(* Release Left Axis *)
IF _SubStep.isActive(2) THEN 
	axis1.Enable:= TRUE;
	IF NOT axis1.State.finish THEN 
		_updateHmiTextWithAxisBusy(axisName:= axisName1);
	ELSIF NOT axis1.State.pass THEN 
		_addressRestart:= _SubStep.actual;
		_subStepError:= "Left axis in error";;
		_subStepMessage:= axis1.State.description;
		_SubStep.set(request:= _SUB_ADDRESS_RETRY_ABORT);
	ELSE 
		_SubStep.INC();
	END_IF
END_IF
(* Reset Axis Right *)
IF _SubStep.isActive(3) THEN 
	IF axis2.Fault THEN 
	axis2.ResetFault();
		IF NOT axis2.AxisError THEN 
			_SubStep.INC();
		ELSE 
			_updateHmiTextWithAxisBusy(axisName:= axisName2); 
		END_IF
	ELSE 
		_SubStep.INC();
	END_IF
END_IF

(* Enable Axis Right *)
IF _SubStep.isActive(4) THEN 
	axis2.Ex_On();
	IF NOT axis2.State.finish THEN 
		_updateHmiTextWithAxisBusy(axisName:= axisName2);
	ELSIF NOT axis2.State.pass THEN 
		_subStepError:= "Right axis in error";
		_subStepMessage:= axis2.State.description;
		_SubStep.set(request:= _SUB_ADDRESS_RETRY_ABORT);
	ELSIF axis2.AxisIsOn THEN 
		_SubStep.INC();
	ELSE 
		_updateHmiTextWithAxisBusy(axisName:= axisName2);
	END_IF
END_IF

(* Release Axis Right *)
IF _SubStep.isActive(5) THEN 
	axis2.Enable:= TRUE;
	IF NOT axis2.State.finish THEN 
		_updateHmiTextWithAxisBusy(axisName:= axisName2);
	ELSIF NOT axis2.State.pass THEN 
		_subStepError:= "Right axis in error";;
		_subStepMessage:= axis2.State.description;
		_SubStep.set(request:= _SUB_ADDRESS_RETRY_ABORT);
	ELSE 
		_SubStep.set(request:= _SUB_ADDRESS_PASS);
	END_IF
END_IF
(* Pass *)
IF _SubStep.isActive(_SUB_ADDRESS_PASS) THEN 
	_step.Condition:= TRUE;
END_IF

(* Fail - Retry/Abort *)
IF _SubStep.isActive(_SUB_ADDRESS_RETRY_ABORT) THEN 
	_retryAbort(
		numOfTargetRetries	:= _UNLIMITED_RETRY_NUMBER,
		retryAddress		:= _addressRestart,
		abortAddress		:= _step.actual);
END_IF

_step.Control();
END_METHOD

METHOD PROTECTED _a2_X_InitAxesToStartProcess
VAR_INPUT
	axis1			: REFERENCE TO KOSTAL_AF2024_Drivers_Actuation_Axis_Festo_CMMT_AS.FB_FESTO_CMMT_AS;
	axisName1		: KOSTAL_AF2024_Core_Settings.T_MaxString;
	axis2			: REFERENCE TO KOSTAL_AF2024_Drivers_Actuation_Axis_Festo_CMMT_AS.FB_FESTO_CMMT_AS;
	axisName2		: KOSTAL_AF2024_Core_Settings.T_MaxString;
END_VAR
(* Reset Axis Left *)
IF _SubStep.isActive(0) THEN 
	IF axis1.Fault THEN 
	axis1.ResetFault();
		IF NOT axis1.Fault THEN 
			_SubStep.INC();
		ELSE 
			_updateHmiTextWithAxisBusy(axisName:= axisName1);
		END_IF
	ELSE 
		_SubStep.INC();
	END_IF
END_IF

(* Reset Axis Right *)
IF _SubStep.isActive(1) THEN 
	IF axis2.Fault THEN 
	axis2.ResetFault();
		IF NOT axis2.Fault THEN 
			_SubStep.INC();
		ELSE 
			_updateHmiTextWithAxisBusy(axisName:= axisName2);
		END_IF
	ELSE 
		_SubStep.INC();
	END_IF
END_IF

(* Enable Axis  Left And Right *)
IF _SubStep.isActive(2) THEN 
	IF axis1.AxisIsOn AND axis2.AxisIsOn THEN 
		_SubStep.INC();
	ELSE 
		axis1.Ex_On();
		axis2.Ex_On();
		IF NOT axis1.State.finish THEN 
			_updateHmiTextWithAxisBusy(axisName:= axisName1);
		ELSIF NOT axis2.State.finish THEN 
			_updateHmiTextWithAxisBusy(axisName:= axisName2);
		ELSIF NOT axis1.State.pass THEN 
			_addressRestart:= _SubStep.actual;
			_getAxisErrorTexts(
				name		:= axisName1,
				description	:= axis1.State.description);
			_SubStep.set(request:= _SUB_ADDRESS_RETRY_ABORT);
		ELSIF NOT axis2.State.pass THEN 
			_addressRestart:= _SubStep.actual;
			_getAxisErrorTexts(
				name		:= axisName2,
				description	:= axis1.State.description);
			_SubStep.set(request:= _SUB_ADDRESS_RETRY_ABORT);
		ELSE 
			_updateHmiTextWithAxisBusy(axisName:= "Both");
		END_IF
	END_IF
END_IF 

(* Release Axes *)
IF _SubStep.isActive(3) THEN 
	axis1.Enable:= TRUE; 
	axis2.Enable:= TRUE; 
	_SubStep.set(request:= _SUB_ADDRESS_PASS);
END_IF

(* Pass *)
IF _SubStep.isActive(_SUB_ADDRESS_PASS) THEN 
	_step.Condition:= TRUE;
END_IF

(* Fail - Retry/Abort *)
IF _SubStep.isActive(_SUB_ADDRESS_RETRY_ABORT) THEN 
	_retryAbort(
		numOfTargetRetries	:= _UNLIMITED_RETRY_NUMBER,
		retryAddress		:= _addressRestart,
		abortAddress		:= _step.actual);
END_IF

_step.Control();
END_METHOD

METHOD PROTECTED _a2_X_InitAxis
VAR_INPUT
	axis			: REFERENCE TO  KOSTAL_AF2024_Drivers_Actuation_Axis_Festo_CMMT_AS.FB_FESTO_CMMT_AS;
	axisName		: KOSTAL_AF2024_Core_Settings.T_MaxString;
END_VAR
(* Reset Axis X *)
IF _SubStep.isActive(0) THEN 
	IF axis.Fault THEN 
	axis.ResetFault();
		IF NOT axis.Fault THEN 
			_SubStep.INC();
		ELSE 
			_updateHmiTextWithAxisBusy(axisName:= axisName);
		END_IF
	ELSE 
		_SubStep.INC();
	END_IF
END_IF

(* Enable Axis *)
IF _SubStep.isActive(1) THEN 
	axis.Ex_On();
	IF NOT axis.State.finish THEN 
		_updateHmiTextWithAxisBusy(axisName:= axisName);
	ELSIF NOT axis.State.pass THEN 
		_addressRestart:= _SubStep.actual;
		_subStepError:= " Axis in error";;
		_subStepMessage:= axis.State.description;
		_SubStep.set(request:= _SUB_ADDRESS_RETRY_ABORT);
	ELSIF axis.AxisIsOn THEN 
		_SubStep.INC();
	ELSE 
		_updateHmiTextWithAxisBusy(axisName:= axisName);
	END_IF
END_IF

(* Release Axis *)
IF _SubStep.isActive(2) THEN 
	axis.Enable:= TRUE;
	IF NOT axis.State.finish THEN 
		_updateHmiTextWithAxisBusy(axisName:= axisName);
	ELSIF NOT axis.State.pass THEN 
		_addressRestart:= _SubStep.actual;
		_subStepError:= "Right axis in errot";;
		_subStepMessage:= axis.State.description;
		_SubStep.set(request:= _SUB_ADDRESS_RETRY_ABORT);
	ELSE 
		_SubStep.set(request:= _SUB_ADDRESS_PASS);
	END_IF
END_IF

(* Pass *)
IF _SubStep.isActive(_SUB_ADDRESS_PASS) THEN 
	_step.Condition:= TRUE;
END_IF

(* Fail - Retry/Abort *)
IF _SubStep.isActive(_SUB_ADDRESS_RETRY_ABORT) THEN 
	_retryAbort(
		numOfTargetRetries	:= _UNLIMITED_RETRY_NUMBER,
		retryAddress		:= _addressRestart,
		abortAddress		:= _step.actual);
END_IF

_step.Control();
END_METHOD

METHOD PROTECTED _a2_X_InitAxisTC3
VAR_INPUT
	axis		: I_LinearAxis_position;
	axisName	: KOSTAL_AF2024_Core_Settings.T_MaxString;
END_VAR
IF _step.toggle THEN 
	_stepDescription:= "InitAxis";
END_IF

(* Reset Axis X *)
IF _SubStep.isActive(0) THEN 
	IF axis.IlinearAxis_Fault THEN 
		axis.IlinearAxis_ResetFault();
		IF NOT axis.IlinearAxis_Fault THEN 
			_SubStep.INC();
		ELSE 
			_updateHmiTextWithAxisBusy(axisName:= axisName);
		END_IF
	ELSE 
		_SubStep.INC();
	END_IF
END_IF

(* Enable Axis *)
IF _SubStep.isActive(1) THEN 
	axis.IlinearAxis_On();
	IF NOT axis.IlinearAxis_State.finish THEN 
		_updateHmiTextWithAxisBusy(axisName:= axisName);
	ELSIF NOT axis.IlinearAxis_State.pass THEN 
		_addressRestart:= _SubStep.actual;
		_getAxisErrorTexts(
			name		:= axisName,
			description	:= STRING_TO_WSTRING(axis.IlinearAxis_State.description));
		_SubStep.set(request:= _SUB_ADDRESS_RETRY_ABORT);
	ELSIF axis.IlinearAxis_isOn THEN 
		_SubStep.INC();
	ELSE 
		_updateHmiTextWithAxisBusy(axisName:= axisName);
	END_IF
END_IF

(* Release Axis *)
IF _SubStep.isActive(2) THEN 
	axis.IlinearAxis_Release(release:= TRUE);
	IF NOT axis.IlinearAxis_State.finish THEN 
		_updateHmiTextWithAxisBusy(axisName:= axisName);
	ELSIF NOT axis.IlinearAxis_State.pass THEN 
		_addressRestart:= _SubStep.actual;
		_getAxisErrorTexts(
			name 			:= axisName,
			description		:= STRING_TO_WSTRING(axis.IlinearAxis_State.description));
		_SubStep.set(request:= _SUB_ADDRESS_RETRY_ABORT);
	ELSE 
		_SubStep.set(request:= _SUB_ADDRESS_PASS);
	END_IF
END_IF

(* Pass *)
IF _SubStep.isActive(_SUB_ADDRESS_PASS) THEN 
	_step.Condition:= TRUE;
END_IF

(* Fail - Retry/Abort *)
IF _SubStep.isActive(_SUB_ADDRESS_RETRY_ABORT) THEN 
	_retryAbort(
		numOfTargetRetries	:= _UNLIMITED_RETRY_NUMBER,
		retryAddress		:= _addressRestart,
		abortAddress		:= _step.actual);
END_IF

_step.Control();
END_METHOD

METHOD PROTECTED _a2_X_InitAxisToStartProcess
VAR_INPUT
	axis			: REFERENCE TO  KOSTAL_AF2024_Drivers_Actuation_Axis_Festo_CMMT_AS.FB_FESTO_CMMT_AS;
	axisName		: KOSTAL_AF2024_Core_Settings.T_MaxString;
END_VAR
(* Reset Axis Left *)
IF _SubStep.isActive(0) THEN 
	IF axis.Fault THEN 
	axis.ResetFault();
		IF NOT axis.Fault THEN 
			_SubStep.INC();
		ELSE 
			_updateHmiTextWithAxisBusy(axisName:= axisName);
		END_IF
	ELSE 
		_SubStep.INC();
	END_IF
END_IF
(* Enable Axis Z *)
IF _SubStep.isActive(1) THEN 
	IF axis.AxisIsOn  THEN 
		_SubStep.INC();
	ELSE 
		axis.Ex_On();
		IF NOT axis.State.finish THEN 
			_updateHmiTextWithAxisBusy(axisName:= axisName);
		ELSIF NOT axis.State.pass THEN 
			_addressRestart:= _SubStep.actual;
			_getAxisErrorTexts(
				name		:= axisName,
				description	:= axis.State.description);
			_SubStep.set(request:= _SUB_ADDRESS_RETRY_ABORT);
		ELSE 
			_updateHmiTextWithAxisBusy(axisName:= axisName);
		END_IF
	END_IF
END_IF 

(* Release Axes *)
IF _SubStep.isActive(2) THEN 
	axis.Enable:= TRUE; 
	_SubStep.set(request:= _SUB_ADDRESS_PASS);
END_IF

(* Pass *)
IF _SubStep.isActive(_SUB_ADDRESS_PASS) THEN 
	_step.Condition:= TRUE;
END_IF

(* Fail - Retry/Abort *)
IF _SubStep.isActive(_SUB_ADDRESS_RETRY_ABORT) THEN 
	_retryAbort(
		numOfTargetRetries	:= _UNLIMITED_RETRY_NUMBER,
		retryAddress		:= _addressRestart,
		abortAddress		:= _step.actual);
END_IF

_step.Control();
END_METHOD

METHOD PROTECTED _a2_X_InitAxisToStartProcessTC3
VAR_INPUT
	axis		: I_LinearAxis_position;
	axisName	: KOSTAL_AF2024_Core_Settings.T_MaxString;
END_VAR
IF _step.toggle THEN 
	_stepDescription:= "InitAxisToStartProcess";
END_IF

(* Reset Axis X *)
IF _SubStep.isActive(0) THEN 
	IF axis.IlinearAxis_Fault THEN 
		axis.IlinearAxis_ResetFault();
		IF NOT axis.IlinearAxis_Fault THEN 
			_SubStep.INC();
		ELSE 
			_updateHmiTextWithAxisBusy(axisName:= axisName);
		END_IF
	ELSE 
		_SubStep.INC();
	END_IF
END_IF

(* Enable Axis *)
IF _SubStep.isActive(1) THEN 
	IF axis.IlinearAxis_isOn THEN 
		_SubStep.INC();
	ELSE 
		axis.IlinearAxis_On();
		IF NOT axis.IlinearAxis_State.finish THEN 
			_updateHmiTextWithAxisBusy(axisName:= axisName);
		ELSIF NOT axis.IlinearAxis_State.pass THEN 
			_addressRestart:= _SubStep.actual;
			_getAxisErrorTexts(
				name		:= axisName,
				description	:= STRING_TO_WSTRING(axis.IlinearAxis_State.description));
			_SubStep.set(request:= _SUB_ADDRESS_RETRY_ABORT);
		ELSE 
			_updateHmiTextWithAxisBusy(axisName:= axisName);
		END_IF
	END_IF
END_IF 

(* Release Axis *)
IF _SubStep.isActive(2) THEN 
	axis.IlinearAxis_Release(release:= TRUE);
	_SubStep.set(request:= _SUB_ADDRESS_PASS);
END_IF

(* Pass *)
IF _SubStep.isActive(_SUB_ADDRESS_PASS) THEN 
	_step.Condition:= TRUE;
END_IF

(* Fail - Retry/Abort *)
IF _SubStep.isActive(_SUB_ADDRESS_RETRY_ABORT) THEN 
	_retryAbort(
		numOfTargetRetries		:= _UNLIMITED_RETRY_NUMBER,
		retryAddress			:= _addressRestart,
		abortAddress			:=	_step.actual);
END_IF

_step.Control();
END_METHOD

METHOD PROTECTED _a2_X_MoveAxesTogether
VAR_INPUT
	axisLeft				: I_Axis;
	axisRight				: I_Axis;
	leftAxisName			: KOSTAL_AF2024_Core_Settings.T_MaxString;
	rightAxisName			: KOSTAL_AF2024_Core_Settings.T_MaxString;
	targetPositionLeftAxis	: REAL;
	targetPositionRightAxis	: REAL;
	axisVelocity 			: REAL;
END_VAR
IF _step.toggle THEN 
	_stepDescription:= "MoveAxis";
END_IF

(* Check actual and target position *)
IF _SubStep.isActive(0) THEN 
	IF _checkIfSamePosition(axisLeft.AxisPositionAct, targetPositionLeftAxis) AND _checkIfSamePosition(axisRight.AxisPositionAct, targetPositionRightAxis) THEN 
		_SubStep.set(request:= _SUB_ADDRESS_PASS);
	ELSE 
		axisLeft.TargetVelocity:= axisVelocity;
		axisLeft.Jerk:= 0;
		axisRight.TargetVelocity:= axisVelocity;
		axisRight.Jerk:= 0;
		_SubStep.INC();
	END_IF
END_IF

(* Move to target position *)
IF _SubStep.isActive(1) THEN 
	_addressRestart:= _SubStep.actual;
	axisLeft.Ex_MoveToPosition(position:= targetPositionLeftAxis);
	axisRight.Ex_MoveToPosition(position:= targetPositionRightAxis);
	IF axisLeft.AxisError THEN 
		_subStepError:= leftAxisName;  
		_subStepMessage:= axisLeft.State.description;
		_SubStep.set(request:= _SUB_ADDRESS_RETRY_ABORT);
	ELSIF axisRight.AxisError THEN 
		_subStepError:= rightAxisName;
		_subStepMessage:= axisRight.State.description;
		_SubStep.set(request:= _SUB_ADDRESS_RETRY_ABORT);
	ELSIF NOT axisLeft.State.finish OR axisLeft.State.busy THEN 
		_updateHmiTextWithAxisBusy(axisName:= leftAxisName);
	ELSIF NOT axisRight.State.finish  THEN 
		_updateHmiTextWithAxisBusy(axisName:= rightAxisName);
	ELSIF NOT axisLeft.State.pass THEN 
		_subStepError:= leftAxisName;
		_subStepMessage:= axisLeft.State.description;
		_SubStep.set(request:= _SUB_ADDRESS_RETRY_ABORT);
	ELSIF NOT axisRight.State.pass THEN 
		_subStepError:= rightAxisName;
		_subStepMessage:= axisLeft.State.description;
		_SubStep.set(request:= _SUB_ADDRESS_RETRY_ABORT);
	ELSE 
		_SubStep.set(request:= _SUB_ADDRESS_PASS);
	END_IF
END_IF

(* Pass *)
IF _SubStep.isActive(_SUB_ADDRESS_PASS) THEN 
	_step.Condition:= TRUE;
END_IF

(* Fail - Retry/Abort *)
IF _SubStep.isActive(_SUB_ADDRESS_RETRY_ABORT) THEN 
	_retryAbort(
		numOfTargetRetries		:= _UNLIMITED_RETRY_NUMBER,
		retryAddress			:= _addressRestart,
		abortAddress			:= _ADDRESS_RUNOUT);
END_IF

_step.Control();
END_METHOD

METHOD PROTECTED _a2_X_MoveAxesTogetherTC3 
VAR_INPUT
	axisLeft				: I_LinearAxis_position;
	axisRight				: I_LinearAxis_position;
	axisName				: KOSTAL_AF2024_Core_Settings.T_MaxString;
	targetPositionLeftAxis	: REAL;
	targetPositionRightAxis	: REAL;
	axisVelocity 			: REAL;
END_VAR
IF _step.toggle THEN 
	_stepDescription:= "MoveAxis";
END_IF

(* Check actual and target position *)
IF _SubStep.isActive(0) THEN 
	IF _checkIfSamePosition(axisLeft.IlinearAxis_PositionAct, targetPositionLeftAxis) AND _checkIfSamePosition(axisRight.IlinearAxis_PositionAct, targetPositionRightAxis) THEN 
		_SubStep.set(request:= _SUB_ADDRESS_PASS);
	ELSE 
		axisLeft.IlinearAxis_Speed:= axisVelocity;
		axisLeft.IlinearAxis_Jerk:= 0;
		axisRight.IlinearAxis_Speed:= axisVelocity;
		axisRight.IlinearAxis_Jerk:= 0;
		_SubStep.INC();
	END_IF
END_IF

(* Move to target position *)
IF _SubStep.isActive(1) THEN 
	_addressRestart:= _SubStep.actual;
	axisLeft.IlinearAxis_MoveToPosition(position:= targetPositionLeftAxis);
	axisRight.IlinearAxis_MoveToPosition(position:= targetPositionRightAxis);
	IF axisLeft.IlinearAxis_Fault THEN 
		_getAxisErrorTexts(
			name		:= "AxisZ-left",
			description	:= STRING_TO_WSTRING(axisLeft.IlinearAxis_State.description));
		_SubStep.set(request:= _SUB_ADDRESS_RETRY_ABORT);
	ELSIF axisRight.IlinearAxis_Fault THEN 
		_getAxisErrorTexts(
			name		:= "AxisZ-right",
			description	:= STRING_TO_WSTRING(axisLeft.IlinearAxis_State.description));
		_SubStep.set(request:= _SUB_ADDRESS_RETRY_ABORT);
	ELSIF NOT axisLeft.IlinearAxis_State.finish OR axisLeft.IlinearAxis_State.busy THEN 
		_updateHmiTextWithAxisBusy(axisName:= axisName);
	ELSIF NOT axisRight.IlinearAxis_State.finish OR axisRight.IlinearAxis_State.busy THEN 
		_updateHmiTextWithAxisBusy(axisName:= axisName);
	ELSIF NOT axisLeft.IlinearAxis_State.pass THEN 
		_getAxisErrorTexts(
			name		:= "AxisZ-left",
			description	:= STRING_TO_WSTRING(axisLeft.IlinearAxis_State.description));
		_SubStep.set(request:= _SUB_ADDRESS_RETRY_ABORT);
	ELSIF NOT axisRight.IlinearAxis_State.pass THEN 
		_getAxisErrorTexts(
			name		:= "AxisZ-right",
			description	:= STRING_TO_WSTRING(axisRight.IlinearAxis_State.description));
		_SubStep.set(request:= _SUB_ADDRESS_RETRY_ABORT);
	ELSE 
		_SubStep.set(request:= _SUB_ADDRESS_PASS);
	END_IF
END_IF

(* Pass *)
IF _SubStep.isActive(_SUB_ADDRESS_PASS) THEN 
	_step.Condition:= TRUE;
END_IF

(* Fail - Retry/Abort *)
IF _SubStep.isActive(_SUB_ADDRESS_RETRY_ABORT) THEN 
	_retryAbort(
		numOfTargetRetries		:= _UNLIMITED_RETRY_NUMBER,
		retryAddress			:= _addressRestart,
		abortAddress			:= _ADDRESS_RUNOUT);
END_IF

_step.Control();
END_METHOD

METHOD PROTECTED _a2_X_MoveAxisToPosition
VAR_INPUT
	axis				: I_Axis;
	axisName			: KOSTAL_AF2024_Core_Settings.T_MaxString;
	targetPosition		: REAL;
	axisVelocity 		: REAL;
END_VAR
IF _step.toggle THEN 
	_stepDescription:= "MoveAxis";
END_IF

(* Check actual and target position *)
IF _SubStep.isActive(0) THEN 
	IF _checkIfSamePosition(actualPosition:= axis.PositionAct, targetPosition:= targetPosition) THEN 
		_SubStep.set(request:= _SUB_ADDRESS_PASS);
	ELSE 
		axis.TargetVelocity:= axisVelocity;
		axis.Jerk:= 0;
		_SubStep.INC();
	END_IF
END_IF

(* Move to target position *)
IF _SubStep.isActive(1) THEN 
	_addressRestart:= _SubStep.actual;
	axis.Ex_MoveToPosition(position:= targetPosition);
	IF axis.AxisError THEN 
		_subStepError:=axisName;
		_subStepMessage:= axis.State.description;
			_SubStep.set(request:= _SUB_ADDRESS_RETRY_ABORT);
	ELSIF NOT axis.State.finish OR axis.State.busy THEN 
		_updateHmiTextWithAxisBusy(axisName:= axisName);
	ELSIF NOT axis.State.pass THEN 
		_subStepError:=axisName;
		_subStepMessage:= axis.State.description;
		_SubStep.set(request:= _SUB_ADDRESS_RETRY_ABORT);
	ELSE 
		_SubStep.set(request:= _SUB_ADDRESS_PASS);
	END_IF
END_IF

(* Pass *)
IF _SubStep.isActive(_SUB_ADDRESS_PASS) THEN 
	_step.Condition:= TRUE;
END_IF

(* Fail - Retry/Abort *)
IF _SubStep.isActive(_SUB_ADDRESS_RETRY_ABORT) THEN 
	_retryAbort(
		numOfTargetRetries		:= _UNLIMITED_RETRY_NUMBER,
		retryAddress			:= _addressRestart,
		abortAddress			:= _ADDRESS_RUNOUT);
END_IF

_step.Control();
END_METHOD

METHOD PROTECTED _a2_X_MoveAxisToPositionTC3 
VAR_INPUT
	axis				: I_LinearAxis_position;

	
	axisName			: KOSTAL_AF2024_Core_Settings.T_MaxString;
	targetPosition		: REAL;
	axisVelocity 		: REAL;
END_VAR
IF _step.toggle THEN 
	_stepDescription:= "MoveAxis";
END_IF

(* Check actual and target position *)
IF _SubStep.isActive(0) THEN 
	IF _checkIfSamePosition(actualPosition:= axis.IlinearAxis_PositionAct, targetPosition:= targetPosition) THEN 
		_SubStep.set(request:= _SUB_ADDRESS_PASS);
	ELSE 
		axis.IlinearAxis_Speed:= axisVelocity;
		axis.IlinearAxis_Jerk:= 0;
		_SubStep.INC();
	END_IF
END_IF

(* Move to target position *)
IF _SubStep.isActive(1) THEN 
	_addressRestart:= _SubStep.actual;
	axis.IlinearAxis_MoveToPosition(position:= targetPosition);
	IF axis.IlinearAxis_Fault THEN 
		_getAxisErrorTexts(
			name		:= axisName,
			description	:= STRING_TO_WSTRING(axis.IlinearAxis_State.description));
			_SubStep.set(request:= _SUB_ADDRESS_RETRY_ABORT);
	ELSIF NOT axis.IlinearAxis_State.finish OR axis.IlinearAxis_State.busy THEN 
		_updateHmiTextWithAxisBusy(axisName:= axisName);
	ELSIF NOT axis.IlinearAxis_State.pass THEN 
		_getAxisErrorTexts(
			name		:= axisName,
			description	:= STRING_TO_WSTRING(axis.IlinearAxis_State.description));
		_SubStep.set(request:= _SUB_ADDRESS_RETRY_ABORT);
	ELSE 
		_SubStep.set(request:= _SUB_ADDRESS_PASS);
	END_IF
END_IF

(* Pass *)
IF _SubStep.isActive(_SUB_ADDRESS_PASS) THEN 
	_step.Condition:= TRUE;
END_IF

(* Fail - Retry/Abort *)
IF _SubStep.isActive(_SUB_ADDRESS_RETRY_ABORT) THEN 
	_retryAbort(
		numOfTargetRetries		:= _UNLIMITED_RETRY_NUMBER,
		retryAddress			:= _addressRestart,
		abortAddress			:= _ADDRESS_RUNOUT);
END_IF

_step.Control();
END_METHOD

METHOD PROTECTED _a2_X_OpenSlider
VAR_INPUT
END_VAR
IF _step.toggle THEN
	_timerSliderInFrontPos(IN:= FALSE);
	_stepDescription:= "OpenSlider";
END_IF

(* If slider in front position skip this step *)
IF _SubStep.isActive(0) THEN
	_timerSliderInFrontPos(IN:= FALSE);
	_addressRestart:= _SubStep.actual;
	IF DI_SliderInFrontPos THEN
		_SubStep.set(request:= 3);
	ELSE
		_SubStep.INC();
	END_IF
END_IF
(* Unlock *)
IF _SubStep.isActive(1) THEN
	IF _SliderLockCylinderInFrontPosition.moveTo_B() THEN
		_SubStep.INC();
	ELSIF _SliderLockCylinderInFrontPosition.Error.active THEN
		_addressRestart:= _SubStep.actual;
		_getCylinderErrorTexts(Cylinder:= _SliderLockCylinderInFrontPosition);
		_SubStep.set(request:= _SUB_ADDRESS_RETRY_ABORT);
	ELSE
		_updateHmiTextWithCylinderTextMoveToHP(Cylinder:= _SliderLockCylinderInFrontPosition);
	END_IF
END_IF
(* Wait slider in back position *)
IF _SubStep.isActive(2) THEN
	_timerSliderInFrontPos(
		IN:= DI_SliderInFrontPos,
		PT:= T#500MS);
	IF NOT DI_SliderInFrontPos THEN
		_Text.ClearVars();
		_Text.AddVar(Text:= _sliderInFrontPositionName);
		_updateHmiText(
			userMessage		:= _Text.GetText(Number:= _E_TextCommon.waitSliderInFrontPosition),
			userAction		:= _Text.GetText(Number:= _E_TextCommon.waitForSensor_0),
			isErrorMessage	:= FALSE);
	ELSIF _timerSliderInFrontPos.Q THEN
		_updateHmiText(
			userMessage		:= _Text.GetText(Number:= _E_TextCommon.waitSliderInFrontPosition),
			userAction		:= _Text.GetText(Number:= _E_TextCommon.waitForSensor_0),
			isErrorMessage	:= FALSE);
	ELSE 
		_SubStep.INC();	
	END_IF
END_IF
(* Lock slider in front position *)
IF _SubStep.isActive(3) THEN
	
	IF _SliderLockCylinderInFrontPosition.moveTo_A() THEN 
		_SubStep.set(request:= _SUB_ADDRESS_PASS);
	ELSIF _SliderLockCylinderInFrontPosition.Error.active THEN
		_getCylinderErrorTexts(Cylinder:= _SliderLockCylinderInFrontPosition);
		_SubStep.set(request:= _SUB_ADDRESS_RETRY_ABORT);
	ELSE
		_updateHmiTextWithCylinderTextMoveToWP(Cylinder:= _SliderLockCylinderInFrontPosition);
	END_IF
END_IF
(* Pass *)
IF _SubStep.isActive(_SUB_ADDRESS_PASS) THEN
	_step.Condition:= TRUE;
END_IF
(* Fail *)
IF _SubStep.isActive(_SUB_ADDRESS_RETRY_ABORT) THEN
	_retryAbort(
		numOfTargetRetries	:= _UNLIMITED_RETRY_NUMBER,
		retryAddress		:= _addressRestart,
		abortAddress		:= _ADDRESS_RUNOUT); 
END_IF

_step.Control();
END_METHOD

METHOD PROTECTED _checkIfSamePosition : BOOL
VAR_INPUT
	actualPosition 			: LREAL;
	targetPosition			: LREAL;
END_VAR
IF (actualPosition >= (targetPosition - 1)) AND (actualPosition <= (targetPosition + 1)) THEN 
	_checkIfSamePosition:= TRUE;
ELSE 
	_checkIfSamePosition:= FALSE;
END_IF
END_METHOD

PROPERTY sliderInBackPositionName : KOSTAL_AF2024_Core_Settings.T_MaxString
GET
sliderInBackPositionName:= _sliderInBackPositionName;
END_GET
SET
_sliderInBackPositionName:= sliderInBackPositionName;
END_SET
END_PROPERTY

PROPERTY sliderInFrontPositionName : KOSTAL_AF2024_Core_Settings.T_MaxString
GET
sliderInFrontPositionName:= _sliderInFrontPositionName;
END_GET
SET
_sliderInFrontPositionName:= sliderInFrontPositionName;
END_SET
END_PROPERTY

END_FUNCTION_BLOCK

// ---- 03_FreeStations/01_Safety/DUTs/T_E_text_Safety.TcPOU
FUNCTION_BLOCK T_E_text_Safety EXTENDS T_E_text_Common
VAR
END_VAR

PROPERTY errorDoor_0 : ST_E_Text
GET
errorDoor_0.Number:= 13;
END_GET
END_PROPERTY

PROPERTY errorEStop_0 : ST_E_Text
GET
errorEStop_0.Number:= 12;
END_GET
END_PROPERTY

PROPERTY errorGroupCom : KOSTAL_AF2024_Core_Text.ST_E_Text
GET
errorGroupCom.Number:= 10;
END_GET
END_PROPERTY

PROPERTY errorGroupFb : ST_E_Text
GET
errorGroupFb.Number:= 11;
END_GET
END_PROPERTY

PROPERTY safetyNok : ST_E_Text
GET
safetyNok.Number:= 5;
END_GET
END_PROPERTY

PROPERTY safetyOk : ST_E_Text
GET
safetyOk.Number:= 4;
END_GET
END_PROPERTY

PROPERTY safetyRelay_0 : ST_E_Text
GET
safetyRelay_0.Number:= 14;
END_GET
END_PROPERTY

END_FUNCTION_BLOCK

// ---- 03_FreeStations/01_Safety/FB_Safety_ST80.TcPOU
FUNCTION_BLOCK FB_Safety_ST80 EXTENDS FB_SafetyBase
VAR
	(* Safety I&O *)
	DI_SafetyRelayInFault 	AT %I* : BOOL;
//	SI_GroupComError	AT %I* : BOOL;
//	SI_GroupFbError		AT %I* : BOOL;
//	SI_SafetyRealyInFault AT %I* : BOOL;
	SI_EstopOk			AT %I* : BOOL;
//	SI_FrontDoorOk		AT %I* : BOOL;
	SO_GroupRun			AT %Q* : BOOL:= TRUE;
//	SO_GroupErrorAck	AT %Q* : BOOL;
//	SO_EStopRestart		AT %Q* : BOOL;
	SO_EStopRestart				: BOOL;
	SO_ResetSafetyExistingSt	AT %Q*	: BOOL; //DO5 20DO1
	SI_FrontDoorOk				: BOOL;
	(* I&O *)
	DO_FrontDoorLock	AT %Q* : BOOL;
	_timerEstopFault	: Tc2_Standard.TON;
	_timerDoorFault		: Tc2_Standard.TON;
END_VAR

METHOD PROTECTED _handleSafety 
VAR_INPUT
END_VAR
_timerEstopFault(
	IN:= NOT SI_EstopOk,
	PT:= T#100MS);
_timerDoorFault(
	IN:= NOT DO_FrontDoorLock,
	PT:= T#100MS);

IF _timerEstopFault.Q THEN
	_Text.ClearVars();
	_Text.AddVar(Text:= "-15S1");
	_message.clear();
	_message.line_01:= _Text.GetText(Number:= _E_Text.errorEStop_0);
	_condition.setMessage(
		priority:= _condition.PriorityLevel_Error,
		message	:= _message);
ELSIF _timerDoorFault.Q THEN
	_Text.ClearVars();
	_Text.AddVar(Text:= "-15S2");
	_message.clear();
	_message.line_01:= _Text.GetText(Number:= _E_Text.errorDoor_0);
	_condition.setMessage(
		priority:= _condition.PriorityLevel_Error,
		message	:= _message);
ELSIF DI_SafetyRelayInFault THEN 
	_Text.ClearVars();
	_Text.AddVar(Text:= "-15U1");
	_message.clear();
	_message.line_01:= "-15U1 Relay in fault";
	_condition.setMessage(
		priority:= _condition.PriorityLevel_Error,
		message	:= _message);
	

END_IF

SO_ResetSafetyExistingSt:= _Hmi_station.Button_Escape.Sign; //HMI restart 
DO_FrontDoorLock:= _doorLock;
_doorLock:= DO_FrontDoorLock;
_isDoorSafe:= DO_FrontDoorLock;
_isDoorUsed:= TRUE;
END_METHOD

END_FUNCTION_BLOCK

// ---- 03_FreeStations/01_Safety/FB_SafetyBase.TcPOU
FUNCTION_BLOCK ABSTRACT FB_SafetyBase EXTENDS KOSTAL_AF2024_Core_Station.FB_Station_Free IMPLEMENTS I_Safety
VAR
	_inHold				: BOOL;
	_isSafe				: BOOL;
	_doorLock			: BOOL;
	_isDoorUsed			: BOOL:= TRUE;
	_isDoorSafe			: BOOL;
	_manual				: BOOL;
	_tempIsSafe			: BOOL;
	_logMessageStart	: BOOL;
	(* Hmi *)
	_Hmi_station		: KOSTAL_AF2024_HMI_WinHMI.FB_Page_Station;
	_E_Text				: T_E_text_Safety;
END_VAR

METHOD PROTECTED ABSTRACT  _handleSafety 
VAR_INPUT
END_VAR
END_METHOD

METHOD PROTECTED _hmiDefine
VAR_INPUT
END_VAR
_Hmi_station.Name:= _Name;

_Hmi_station.Text.line_01:= _condition.Message.line_01;
_Hmi_station.Text.line_02:= _condition.Message.line_02;
_Hmi_station.Text.line_03:= _condition.Message.line_03;

_Hmi_station.Button_Escape.Visible:= (_condition.isError() OR _Hmi_station.Button_Escape.Sign) AND _manual;
_Hmi_station.Button_Escape.Text:= _Text.GetText(Number:= _E_Text.reset);

_Hmi_station.Status.CopyFrom(IN:= _condition);

_Hmi_station.FBmain();
END_METHOD

METHOD PROTECTED _logStart
VAR_INPUT
END_VAR
IF _logMessageStart AND _Text.State.ready AND (_Text.LoadedLanguage <> '') THEN
	IF _log("===START===") THEN
		_logMessageStart:= FALSE;
	END_IF
	
	IF _tempIsSafe THEN 
		_log(Text:= _Text.GetText(Number:= _E_Text.safetyOk));
	ELSE
		_log(Text:= _Text.GetText(Number:= _E_Text.safetyNok));
	END_IF
END_IF
END_METHOD

METHOD PROTECTED _resetCondition 
VAR_INPUT
END_VAR
IF _condition.isError() THEN
	IF _Hmi_station.Button_Escape.Pulse THEN
		_condition.clear();
	END_IF
ELSE
	_condition.clear();
END_IF
END_METHOD

PROPERTY PUBLIC doorLock : BOOL
GET
doorLock:= _doorLock;
END_GET
SET
_doorLock:= doorLock;
END_SET
END_PROPERTY

METHOD FB_init : BOOL
VAR_INPUT
	bInitRetains : BOOL; // if TRUE, the retain variables are initialized (warm start / cold start)
	bInCopyCode : BOOL;  // if TRUE, the instance afterwards gets moved into the copy code (online change)
	ID_Name			: KOSTAL_AF2024_Core_Settings.T_MaxString;
	ID_Key			: DINT;
	CommonText		: KOSTAL_AF2024_Core_Text.I_Text;
	textPath		: KOSTAL_AF2024_Core_Settings.T_MaxString_UTF8;
END_VAR
_TextPath:= textPath;
END_METHOD

METHOD PUBLIC FBmain
VAR_INPUT
END_VAR
IF NOT _parameterControl() THEN RETURN; END_IF
 
_hmiDefine();

IF NOT _TextReader() THEN RETURN; END_IF;

_logStart();
_handleSafety();
_resetCondition();
_tempIsSafe:= NOT _condition.isError();

(* Log if safety state changed *)
IF _isSafe <> _tempIsSafe THEN
	IF _tempIsSafe THEN			
		_log(_Text.GetText(_E_text.safetyOk));
	ELSE							
		_log(_condition.Message.toString());				
	END_IF
END_IF

_isSafe:= _tempIsSafe;

IF _isSafe THEN	
	_message.clear();
	_message.line_01:= _Text.GetText(Number:= _E_text.safetyOk);
	_condition.setMessage(
		priority:= _condition.PriorityLevel_Info, 
		message	:= _message);
END_IF
END_METHOD

PROPERTY inHold : BOOL
GET
inHold:= _inHold;
END_GET
END_PROPERTY

PROPERTY isDoorSafe : BOOL
GET
isDoorSafe:= _isDoorSafe;
END_GET
END_PROPERTY

PROPERTY isDoorUsed : BOOL
GET
isDoorUsed:= _isDoorUsed;
END_GET
END_PROPERTY

PROPERTY isSafe : BOOL
GET
isSafe:= _isSafe;
END_GET
END_PROPERTY

PROPERTY PUBLIC manual : BOOL
GET
manual := _manual;
END_GET
SET
_manual:= manual;
END_SET
END_PROPERTY

END_FUNCTION_BLOCK

// ---- 03_FreeStations/01_Safety/FB_Safety_STAudi.TcPOU
FUNCTION_BLOCK FB_Safety_STAudi EXTENDS FB_SafetyBase
VAR
	(* Safety I&O *)
//	SI_GroupComError	AT %I* : BOOL;
//	SI_GroupFbError		AT %I* : BOOL;
//	SI_SafetyRealyInFault 			AT %I* : BOOL;
//	SO_RunSafety		AT %Q* : BOOL;
//	SO_ErrorAckSafety	AT %Q* : BOOL;
//	SO_ResetSafetyExistingSt		AT %Q* : BOOL;//DO5 20DO1
	SI_EstopOk			AT %I* : BOOL;
	SI_FrontDoorOk		AT %I* : BOOL;
	SI_BackDoorOk		AT %I* : BOOL;
	SO_GroupRun						AT %Q* : BOOL:= TRUE;
//	SO_GroupErrorAck	AT %Q* : BOOL;
//	SO_EStopRestart		AT %Q* : BOOL;
	SO_RestartSaferyRelay		AT %Q* 				   : BOOL; 
//	SI_FrontDoorOk						   : BOOL;
//	SI_BackDoorOk						   : BOOL;
	(* I&O *)
	DO_FrontDoorLock				AT %Q* : BOOL;
	DO_BackDoorLock					AT %Q* : BOOL;
	_timerEstopFault					   : Tc2_Standard.TON;
	_timerFrontDoorFault				   : Tc2_Standard.TON;
	_timerBackDoorFault					   : Tc2_Standard.TON;
END_VAR

METHOD PROTECTED _handleSafety 
VAR_INPUT
END_VAR
_timerEstopFault(
	IN:= NOT SI_EstopOk,
	PT:= T#100MS);
_timerFrontDoorFault(
	IN:= SI_FrontDoorOk,
	PT:= T#100MS);
_timerBackDoorFault(
	IN:= SI_BackDoorOk,
	PT:= T#100MS);

IF _timerEstopFault.Q THEN
	_Text.ClearVars();
	_Text.AddVar(Text:= "11SA1");
	_message.clear();
	_message.line_01:= _Text.GetText(Number:= _E_Text.errorEStop_0);
	_condition.setMessage(
		priority:= _condition.PriorityLevel_Error,
		message	:= _message);
ELSIF _timerFrontDoorFault.Q THEN
	_Text.ClearVars();
	_Text.AddVar(Text:= "11SQ1");
	_message.clear();
	_message.line_01:= _Text.GetText(Number:= _E_Text.errorDoor_0);
	_condition.setMessage(
		priority:= _condition.PriorityLevel_Error,
		message	:= _message);
ELSIF _timerBackDoorFault.Q THEN
	_Text.ClearVars();
	_Text.AddVar(Text:= "11SQ2");
	_message.clear();
	_message.line_01:= _Text.GetText(Number:= _E_Text.errorDoor_0);
	_condition.setMessage(
		priority:= _condition.PriorityLevel_Error,
		message	:= _message);
END_IF

SO_RestartSaferyRelay:= _Hmi_station.Button_Escape.Sign; //HMI restart 
DO_FrontDoorLock:= _doorLock;
DO_BackDoorLock:= _doorLock;
_isDoorSafe:= DO_BackDoorLock AND DO_FrontDoorLock;
_isDoorUsed:= TRUE;
END_METHOD

END_FUNCTION_BLOCK

// ---- 03_FreeStations/01_Safety/FB_Safety_ST50.TcPOU
FUNCTION_BLOCK FB_Safety_ST50 EXTENDS FB_SafetyBase
VAR
	(* Safety I&O *)
//	SI_GroupComError	AT %I* : BOOL;
//	SI_GroupFbError		AT %I* : BOOL;
//	SI_SafetyRealyInFault 			AT %I* : BOOL;
//	SO_RunSafety		AT %Q* : BOOL;
//	SO_ErrorAckSafety	AT %Q* : BOOL;
//	SO_ResetSafetyExistingSt		AT %Q* : BOOL;//DO5 20DO1
	SI_EstopOk			AT %I* : BOOL;
	SI_FrontDoorOk		AT %I* : BOOL;
	SI_BackDoorOk		AT %I* : BOOL;
	SO_GroupRun						AT %Q* : BOOL:= TRUE;
//	SO_GroupErrorAck	AT %Q* : BOOL;
//	SO_EStopRestart		AT %Q* : BOOL;
	SO_RestartSaferyRelay		AT %Q* 				   : BOOL; 
//	SI_FrontDoorOk						   : BOOL;
//	SI_BackDoorOk						   : BOOL;
	(* I&O *)
	DO_FrontDoorLock				AT %Q* : BOOL;
	DO_BackDoorLock					AT %Q* : BOOL;
	_timerEstopFault					   : Tc2_Standard.TON;
	_timerFrontDoorFault				   : Tc2_Standard.TON;
	_timerBackDoorFault					   : Tc2_Standard.TON;
END_VAR

METHOD PROTECTED _handleSafety 
VAR_INPUT
END_VAR
//_eStop();


_timerEstopFault(
	IN:=  SI_EstopOk, //AND NOT SO_RestartSaferyRelay,
	PT:= T#100MS);
_timerFrontDoorFault(
	IN:= SI_FrontDoorOk,
	PT:= T#100MS);
_timerBackDoorFault(
	IN:= SI_BackDoorOk,
	PT:= T#100MS);


//IF SI_GroupComError THEN
//	_message.clear();
//	_message.line_01:= _Text.GetText(Number:= _E_Text.errorGroupCom);
//	_condition.setMessage(
//		priority:= _condition.PriorityLevel_Error,
//		message	:= _message);
IF _timerEstopFault.Q THEN
	_Text.ClearVars();
	_Text.AddVar(Text:= "11SA1"); //Check Eplan
	_message.clear();
	_message.line_01:= _Text.GetText(Number:= _E_Text.errorEStop_0);
	_condition.setMessage(
		priority:= _condition.PriorityLevel_Error,
		message	:= _message);
ELSIF _timerFrontDoorFault.Q THEN
	_Text.ClearVars();
	_Text.AddVar(Text:= "11SQ1");
	_message.clear();
	_message.line_01:= _Text.GetText(Number:= _E_Text.errorDoor_0);
	_condition.setMessage(
		priority:= _condition.PriorityLevel_Error,
		message	:= _message);
ELSIF _timerBackDoorFault.Q THEN
	_Text.ClearVars();
	_Text.AddVar(Text:= "11SQ2");
	_message.clear();
	_message.line_01:= _Text.GetText(Number:= _E_Text.errorDoor_0);
	_condition.setMessage(
		priority:= _condition.PriorityLevel_Error,
		message	:= _message);
	
	
//ELSIF SI_GroupFbError THEN
//	_message.clear();
//	_message.line_01:= _Text.GetText(Number:= _E_Text.errorGroupFb);
//	_condition.setMessage(
//		priority:= _condition.PriorityLevel_Error,
//		message	:= _message);
END_IF

//SO_RunSafety:= TRUE;
//SO_ErrorAckSafety:= _Hmi_station.Button_Escape.Sign;
//SO_ResetSafetyExistingSt:= SO_ErrorAckSafety; //Da se proveri dali ova vaka kje raboti 
SO_RestartSaferyRelay:= _Hmi_station.Button_Escape.Sign; //HMI restart 
DO_FrontDoorLock:= _doorLock;
DO_BackDoorLock:= _doorLock;
//_doorLock:= SI_FrontDoorOk;
_isDoorSafe:= DO_BackDoorLock AND DO_FrontDoorLock;
_isDoorUsed:= TRUE;
END_METHOD

END_FUNCTION_BLOCK

// ---- 03_FreeStations/02_Parameters/FB_ParameterHandler.TcPOU
FUNCTION_BLOCK FB_ParameterHandler EXTENDS KOSTAL_AF2024_HMI_WinHMI.FB_Parameters_Base IMPLEMENTS I_Parameters_MainControl
VAR
END_VAR

PROPERTY airPressureMax : INT
GET
airPressureMax:= STRING_TO_INT(_getParameterValue(index:= E_Parameters.airPressureMax));
END_GET
END_PROPERTY

PROPERTY airPressureMin : INT
GET
airPressureMin:= STRING_TO_INT(_getParameterValue(index:= E_Parameters.airPressureMin));
END_GET
END_PROPERTY

{warning 'add property implementation'}
PROPERTY cylinderSensorTimeout : TIME
GET
cylinderSensorTimeout:= STRING_TO_TIME(_getParameterValue(index:= E_Parameters.cylinderTimeout));
END_GET
END_PROPERTY

METHOD FB_init : BOOL
VAR_INPUT
	bInitRetains 	: BOOL; // if TRUE, the retain variables are initialized (warm start / cold start)
	bInCopyCode 	: BOOL;  // if TRUE, the instance afterwards gets moved into the copy code (online change)
	ID_Name			: KOSTAL_AF2024_Core_Settings.T_MaxString;
	ID_Key			: DINT;
	CommonText		: KOSTAL_AF2024_Core_Text.I_Text;
	parameterPath	: KOSTAL_AF2024_Core_Settings.T_MaxString_UTF8;
	SystemTime		: KOSTAL_AF2024_Core_GetSystemTime.I_TimeSource;
END_VAR
_fullQualifiedFile:= parameterPath;
_I_getTime:= SystemTime;
END_METHOD

{warning 'add property implementation'}
PROPERTY isLoggerEnabled : BOOL
GET
isLoggerEnabled:= STRING_TO_BOOL(_getParameterValue(index:= E_Parameters.isLoggerEnabled));
END_GET
END_PROPERTY

{warning 'add property implementation'}
PROPERTY isNagaraEnable : BOOL
GET
isNagaraEnable:= STRING_TO_BOOL(_getParameterValue(index:= E_Parameters.isNagaraEnable));
END_GET
END_PROPERTY

{warning 'add property implementation'}
PROPERTY numberOfRetries : INT
GET
airPressureMax:= STRING_TO_INT(_getParameterValue(index:= E_Parameters.numberOfRetries));
END_GET
END_PROPERTY

END_FUNCTION_BLOCK

// ---- 03_FreeStations/03_TextMaster/FB_TextMaster.TcPOU
FUNCTION_BLOCK FB_TextMaster EXTENDS KOSTAL_AF2024_Templates_TextMaster.FB_TextMaster
VAR
	_Hmi_station				: KOSTAL_AF2024_HMI_WinHMI.FB_Page_Station;
END_VAR

METHOD PROTECTED _linkHmi
VAR_INPUT
END_VAR
_iHmi_station := _Hmi_station;
_Hmi_station.FBmain();
END_METHOD

METHOD FB_init : BOOL
VAR_INPUT
	bInitRetains 		: BOOL; // if TRUE, the retain variables are initialized (warm start / cold start)
	bInCopyCode			: BOOL;  // if TRUE, the instance afterwards gets moved into the copy code (online change)
	ID_Name				: KOSTAL_AF2024_Core_Settings.T_MaxString;
	ID_Key				: DINT;
	commonTextPath		: KOSTAL_AF2024_Core_Settings.T_MaxString_UTF8;
	textPath			: KOSTAL_AF2024_Core_Settings.T_MaxString_UTF8;
END_VAR
_pathCommon:= commonTextPath;
_TextPath:= textPath;
END_METHOD

END_FUNCTION_BLOCK

// ---- 03_FreeStations/04_EtherCAT Monitoring/DUTs/T_E_text_EtherCAT.TcPOU
FUNCTION_BLOCK T_E_text_EtherCAT EXTENDS T_E_text_Common
VAR
END_VAR

PROPERTY allDevicesOk : KOSTAL_AF2024_Core_Text.ST_E_Text
GET
allDevicesOk.Number:= 11;
END_GET
END_PROPERTY

PROPERTY device_0_isInState_1 : KOSTAL_AF2024_Core_Text.ST_E_Text
GET
device_0_isInState_1.Number:= 10;
END_GET
END_PROPERTY

PROPERTY name : KOSTAL_AF2024_Core_Text.ST_E_Text
GET
name.Number:= 2;
END_GET
END_PROPERTY

END_FUNCTION_BLOCK

// ---- 03_FreeStations/04_EtherCAT Monitoring/FB_EtherCAT_Base.TcPOU
FUNCTION_BLOCK ABSTRACT FB_EtherCAT_Base EXTENDS KOSTAL_AF2024_Core_Station.FB_Station_Free IMPLEMENTS I_EtherCAT
VAR
	_Hmi_station			: KOSTAL_AF2024_HMI_WinHMI.FB_Page_Station;
	_E_Text					: T_E_text_EtherCAT;
	_inError				: BOOL;
END_VAR

METHOD PROTECTED ABSTRACT _checkAllDevices
VAR_INPUT
END_VAR
END_METHOD

METHOD PROTECTED _hmiDefine
VAR_INPUT
END_VAR
_Hmi_station.FBmain();

_Hmi_station.Name:= _Text.GetText(Number:= _E_Text.name);

_Hmi_station.Text.line_01:= _Hmi_station.Status.Message.line_01;
_Hmi_station.Text.line_02:= _Hmi_station.Status.Message.line_02;
_Hmi_station.Text.line_03:= _Hmi_station.Status.Message.line_03;
(* Reset button *)
_Hmi_station.Button_Escape.Text:= _Text.GetText(Number:= _E_Text.reset);
_Hmi_station.Button_Escape.Visible:= _Hmi_station.Status.isError();

_Hmi_station.Status.CopyFrom(IN:= _condition);
END_METHOD

METHOD PROTECTED _isDeviceOk : BOOL
VAR_INPUT
	state		: INT;
	name		: WSTRING;
END_VAR
IF (state = 8) THEN
	_isDeviceOk:= TRUE;
ELSE
	_Text.ClearVars();
	_Text.AddVar(Text:= name);
	_Text.AddVar(Text:= _stateToString(state:= state));
	_message.clear();
	_message.line_01:= _Text.GetText(Number:= _E_Text.device_0_isInState_1);
	_condition.setMessage(
		priority:= _condition.PriorityLevel_Error,
		message	:= _message);
	_isDeviceOk:= FALSE;
	_inError:= TRUE;
END_IF
END_METHOD

METHOD PROTECTED _resetCondition 
VAR_INPUT
END_VAR
IF _condition.isError() THEN 
	IF _Hmi_station.Button_Escape.Pulse THEN 
		_condition.clear();
	END_IF
ELSE 
	_condition.clear();
END_IF
END_METHOD

METHOD PROTECTED _stateToString : KOSTAL_AF2024_Core_Settings.T_MaxString
VAR_INPUT
	state		: INT;
END_VAR
CASE state OF 
	1: _stateToString := "INIT";
	2: _stateToString := "PREOP";
	3: _stateToString := "BOOT";
	4: _stateToString := "SAFEOP";
	8: _stateToString := "OP";
ELSE 
	_stateToString := "Unknown";
END_CASE
END_METHOD

METHOD FB_init : BOOL
VAR_INPUT
	bInitRetains 	: BOOL; // if TRUE, the retain variables are initialized (warm start / cold start)
	bInCopyCode		: BOOL;  // if TRUE, the instance afterwards gets moved into the copy code (online change)
	ID_Name			: KOSTAL_AF2024_Core_Settings.T_MaxString;
	ID_Key			: DINT;
	CommonText		: KOSTAL_AF2024_Core_Text.I_Text;
	textPath		: KOSTAL_AF2024_Core_Settings.T_MaxString_UTF8;
END_VAR
_textPath:= textPath;
END_METHOD

METHOD FBmain
VAR_INPUT
END_VAR
IF NOT _parameterControl() THEN RETURN; END_IF

_hmiDefine();
_resetCondition();

IF NOT _TextReader() THEN RETURN; END_IF

_inError:= FALSE;
_checkAllDevices();
END_METHOD

PROPERTY inError : BOOL
GET
inError:= _inError;
END_GET
END_PROPERTY

END_FUNCTION_BLOCK

// ---- 03_FreeStations/05_Fuse Monitorning/DUTs/T_E_text_Fuse.TcPOU
FUNCTION_BLOCK T_E_text_Fuse EXTENDS T_E_text_Common
VAR
END_VAR

PROPERTY allFusesOk : KOSTAL_AF2024_Core_Text.ST_E_Text
GET
allFusesOk.Number:= 11;
END_GET
END_PROPERTY

PROPERTY fuse_0_tripped : KOSTAL_AF2024_Core_Text.ST_E_Text
GET
fuse_0_tripped.Number:= 10;
END_GET
END_PROPERTY

PROPERTY name : KOSTAL_AF2024_Core_Text.ST_E_Text
GET
name.Number:= 2;
END_GET
END_PROPERTY

END_FUNCTION_BLOCK

// ---- 03_FreeStations/05_Fuse Monitorning/FB_FuseMonitoringBase.TcPOU
FUNCTION_BLOCK ABSTRACT FB_FuseMonitoringBase EXTENDS KOSTAL_AF2024_Core_Station.FB_Station_Free IMPLEMENTS I_Fuse
VAR
	_Hmi_station			: KOSTAL_AF2024_HMI_WinHMI.FB_Page_Station;
	_E_Text					: T_E_text_Fuse;
	_inError				: BOOL;
END_VAR

METHOD PROTECTED ABSTRACT _checkAllDevices
VAR_INPUT
END_VAR
END_METHOD

METHOD PROTECTED _hmiDefine
VAR_INPUT
END_VAR
_Hmi_station.FBmain();

_Hmi_station.Name:= _Text.GetText(Number:= _E_Text.name);

_Hmi_station.Text.line_01:= _Hmi_station.Status.Message.line_01;
_Hmi_station.Text.line_02:= _Hmi_station.Status.Message.line_02;
_Hmi_station.Text.line_03:= _Hmi_station.Status.Message.line_03;
(* Reset button *)
_Hmi_station.Button_Escape.Text:= _Text.GetText(Number:= _E_Text.reset);
_Hmi_station.Button_Escape.Visible:= _Hmi_station.Status.isError();

_Hmi_station.Status.CopyFrom(IN:= _condition);
END_METHOD

METHOD PROTECTED _resetCondition
VAR_INPUT
END_VAR
IF _condition.isError() THEN
	IF _Hmi_station.Button_Escape.Pulse THEN
		_condition.clear();
	END_IF
ELSE
	_condition.clear();
END_IF
END_METHOD

METHOD FB_init : BOOL
VAR_INPUT
	bInitRetains : BOOL; // if TRUE, the retain variables are initialized (warm start / cold start)
	bInCopyCode : BOOL;  // if TRUE, the instance afterwards gets moved into the copy code (online change)
	ID_Name			: KOSTAL_AF2024_Core_Settings.T_MaxString;
	ID_Key			: DINT;
	CommonText		: KOSTAL_AF2024_Core_Text.I_Text;
	textPath		: KOSTAL_AF2024_Core_Settings.T_MaxString_UTF8;
END_VAR
_textPath:= textPath;
END_METHOD

METHOD PUBLIC FBmain
VAR_INPUT
END_VAR
IF NOT _parameterControl() THEN RETURN; END_IF

_hmiDefine();
_resetCondition();

IF NOT _TextReader() THEN RETURN; END_IF

_inError:= FALSE;
_checkAllDevices();
END_METHOD

PROPERTY inError : BOOL
GET
inError:= _inError;
END_GET
END_PROPERTY

END_FUNCTION_BLOCK

// ---- 04_ComponentSource/FB_CounterHandler.TcPOU
FUNCTION_BLOCK FB_CounterHandler EXTENDS KOSTAL_AF2024_HMI_WinHMI.FB_Counter
VAR
	_scrap				: REAL;
	_FormatString		: Tc2_Utilities.FB_FormatString;
	_FormattedString	: STRING(255);
END_VAR

METHOD PROTECTED _storage
VAR_INPUT
END_VAR


IF	_Istorage.State.fail THEN

	_message.clear();
	_message.line_01:= "ERROR Counter Storage";
	_message.line_02:= _Istorage.State.description;

	_condition.setMessage(_condition.PriorityLevel_Error, _message);
	
	IF _pageStation.Button_Escape.Pulse THEN
		 _Istorage.Reset();
	END_IF

ELSIF NOT _Istorage.State.ready THEN

	_message.clear();
	_message.line_01:= "wait for Counter Storage >Ready<";
	_message.line_02:= _Istorage.State.description;
	
	_condition.setMessage(_condition.PriorityLevel_Message, _message);


ELSIF NOT _initFromStorageDone THEN

	_counterPass.Init(_Istorage.Content.Pass);
	_counterFail.Init(_Istorage.Content.Fail);
	
	_initFromStorageDone:= TRUE;
	
ELSE	
	_Istorage.Content.fail:= _counterFail.Counter;
	_Istorage.Content.Pass:= _counterPass.Counter;
	
	IF (_counterPass.Counter + _counterFail.Counter) > 0 THEN
		_scrap:= UDINT_TO_REAL(_counterFail.Counter)/UDINT_TO_REAL(_counterPass.Counter + _counterFail.Counter)*100;
	ELSE
		_scrap:= 0;
	END_IF
	
	_message.clear();
	_message.line_01:= Tc2_Standard.WCONCAT(
		STR1:= "OK: ",
		STR2:= UDINT_TO_WSTRING(_counterPass.Counter));
	_message.line_02:= Tc2_Standard.WCONCAT(
		STR1:= "NOK: ",
		STR2:= UDINT_TO_WSTRING(_counterFail.Counter));
	_FormatString(
		sFormat:= '%.2f', 
		arg1:= Tc2_Utilities.F_REAL(_scrap), 
		sOut=> _FormattedString);		
	_message.line_03:= Tc2_Standard.WCONCAT(
		STR1:= "Scrap: ",
		STR2:= STRING_TO_WSTRING(_FormattedString));
	_message.line_03:= Tc2_Standard.WCONCAT(
		STR1:= _message.line_03,
		STR2:= "%");
	_condition.setMessage(
		priority:= _condition.PriorityLevel_Text, 
		message	:= _message);
		
	IF _Hmi_station.Button_OnOff.Pulse THEN
		_counterFail.Reset();
		_counterPass.Reset();
	END_IF
END_IF
END_METHOD

END_FUNCTION_BLOCK

// ---- MAIN.TcPOU
PROGRAM MAIN
VAR
	fb : FB_MainControlCell; 
	fb1 : FB_StationBase;
END_VAR

END_PROGRAM
